// TIA Portal V21 export
// export: Created 2026-11-11T00:47:23.0969325Z, ExportSetting WithDefaults, DisplayName Totally Integrated Automation Portal, DisplayVersion V21 Update 3, DisplayName STEP 7 Professional, DisplayVersion V21 Update 3, DisplayName STEP 7 Safety, DisplayVersion V21, DisplayName Tech WebApplication, DisplayVersion V21, DisplayName WinCC Basic/Comfort/Advanced, DisplayVersion V21 Update 3, DisplayName WinCC Unified, DisplayVersion V21 Update 3
FUNCTION_BLOCK "FB_Fbd_ex087"   // FB103, FBD
{ S7_Optimized_Access := 'TRUE' }
VERSION : 0.1
// stored: AutoNumber true, IsIECCheckEnabled false, IsRetainMemResEnabled false, MemoryReserve 100, SetENOAutomatically false, UDAEnableTagReadback false
   VAR_INPUT
      v_pe_i_dev_new : Bool;
      v_error_code : Byte;
   END_VAR
   VAR_OUTPUT
      v_error : Bool;
      v_status : Word;
   END_VAR
   VAR_IN_OUT
      v_activate : Bool;
      v_valid : Bool;
      v_data_errorrsp : Variant;
   END_VAR
BEGIN

REGION Network 1: PE_Error_RSP - Generate negative answer to command
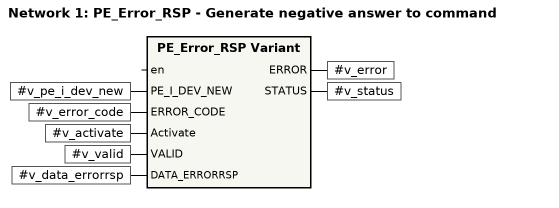
   PE_Error_RSP(PE_I_DEV_NEW := #v_pe_i_dev_new,
                ERROR_CODE := #v_error_code,
                Activate := #v_activate,
                VALID := #v_valid,
                DATA_ERRORRSP := #v_data_errorrsp,
                ERROR => #v_error,
                STATUS => #v_status);
END_REGION
END_FUNCTION_BLOCK
